(* IEC 61131-3 sources: nautilus/lang/conformance/fb-ton, 1 file *)

(* ---- fb-ton.st ---- *)
PROGRAM TonSt
(* TON in Structured Text: the reference path. *)
VAR_EXTERNAL
    IN    : BOOL;
    PT    : TIME;
    st_Q  : BOOL;
    st_ET : TIME;
END_VAR
VAR
    t : TON;
END_VAR

t(IN := IN, PT := PT);
st_Q  := t.Q;
st_ET := t.ET;
END_PROGRAM
